(* IEC 61131-3 sources: Lasal-MCP/examples/SampleSource/LASALScreenAdvancedSolution/LASALScreenAdvancedSolution/LASALScreenAdvacnedSolution/Stations/Terminal/HMI/Network/ScrollNet, 1 file *)

(* ---- ONE_ScrollNet_Table.st ---- *)
#define OBJECTS_CONFIG

FUNCTION GLOBAL TAB ONE_ScrollNet
-1$UINT, 0$UINT,
0$UINT, 0$UINT,

5$UDINT,
TO_UDINT(2980745877), "_MyIO", 0$UINT, 3$UINT, 0$UINT,
TO_UDINT(3043040051), "_ScrollArea", 0$UINT, 15$UINT, 0$UINT,
TO_UDINT(2779823616), "_ScrollArea2", 0$UINT, 8$UINT, 0$UINT,
TO_UDINT(1321167573), "MyHeader", 0$UINT, 0$UINT, 1$UINT,
TO_UDINT(1880544669), "MyScrollList", 0$UINT, 0$UINT, 1$UINT,

_NO_ATTR, TO_UDINT(1965782662), "MYHEADER1",

_NO_ATTR, TO_UDINT(219289243), "MYSCROLLLIST1",

//Internal connections
0$UDINT,
0$UDINT,
0$UDINT,
0$UDINT,

//Initialization values
0$UDINT,
5$UDINT,
TO_UDINT(0), "LineWidth", TO_UDINT(500),//|ScrollNet.MyHeader1.LineWidth;
TO_UDINT(0), "ExtendedScrollBar", TO_UDINT(0),//|ScrollNet.MyHeader1.ExtendedScrollBar;
TO_UDINT(1), "VerticalLevel", TO_UDINT(1),//|ScrollNet.MyScrollList1.VerticalLevel;
TO_UDINT(1), "LineWidth", TO_UDINT(500),//|ScrollNet.MyScrollList1.LineWidth;
TO_UDINT(1), "ExtendedScrollBar", TO_UDINT(0),//|ScrollNet.MyScrollList1.ExtendedScrollBar;

//Symbolic initialization values
0$UDINT,
0$UDINT,

//Initialization of string values
0$UDINT,
0$UDINT,

//Configuration of tasks (RealTime, Cyclic, Background)
0$UDINT,
0$UDINT,

0$UDINT,
0$UDINT,

0$UDINT,
0$UDINT,

//External connections
0$UDINT,
2$UDINT,
TO_UDINT(0), "Lse", C_DIR, TO_UDINT(299963966), "Lse","Lse",
TO_UDINT(1), "Lse", C_DIR, TO_UDINT(299963966), "Lse","Lse",

//Magic internal connections
0$UDINT,
0$UDINT,

//Configuration of timeslots of tasks (RealTime, Cyclic)
#ifdef __LSLLDR_TIMESLOTS__
0$UDINT,
0$UDINT,

0$UDINT,
0$UDINT,

#endif //__LSLLDR_TIMESLOTS__

//MultiMaster connections
#ifdef __LSLLDR_MULTIMASTER__
0$UDINT,
0$UDINT,
#endif //__LSLLDR_MULTIMASTER__

//Configuration for task ID (RealTime, CyclicTime)
#ifdef __LSLLDR_TASKID__
"\\\\TASKS2  "
0$UDINT,
0$UDINT,

0$UDINT,
0$UDINT,

0$UDINT,
0$UDINT,

#endif //__LSLLDR_TASKID__

END_FUNCTION
